(* IEC 61131-3 sources: 2026_Projet_YGO_ExcavatriceDragage/CODE/SIMULATION/PLC_TESTS, 3 files *)

(* ---- GVL_PLC_Tests.st ---- *)
(* ═══════════════════════════════════════════════════════════════
   🧪 GVL_PLC_Tests — Variables globales du banc de validation
   ───────────────────────────────────────────────────────────────
   🎯 Rôle : Regroupe toutes les commandes et retours d'états
      du banc de tests automatique in-PLC.
   ═══════════════════════════════════════════════════════════════ *)

{attribute 'qualified_only'}
VAR_GLOBAL
    CmdRunTests                : BOOL := FALSE; // 🔑 Lancement des tests de validation (bouton IHM/Simu)
    TestInProgress             : BOOL;          // Test en cours d'exécution
    AllTestsPassed             : BOOL;          // Succès global : tous les scénarios validés 🟢
    TestFailed                 : BOOL;          // Échec détecté 🔴
    TC01_NominalArming_Ok      : BOOL;          // Statut TC-01 (Armement nominal & AU)
    TC02_RedundancyFault_Ok    : BOOL;          // Statut TC-02 (Contacteur collé)
    TC03_Lockout_Ok            : BOOL;          // Statut TC-03 (Lockout 5s)
    FailedTestCase             : INT;           // Index du scénario en échec

    // Signaux de surcharge internes (pilotés par le validateur de test)
    OverrideChainTrue          : BOOL;          // Force la boucle AU à TRUE
    OverrideChainFalse         : BOOL;          // Force la boucle AU à FALSE
    OverrideContactorFalse     : BOOL;          // Force le retour contacteur à FALSE
END_VAR

(* ---- FB_PLC_Tests_Management.st ---- *)
(* ═══════════════════════════════════════════════════════════════
   🧪 FB_PLC_Tests_Management — Gestion Globale des Tests de Validation Automatisés
   ───────────────────────────────────────────────────────────────
   🎯 Rôle : Regroupe, configure et orchestre toutes les instances
      de tests de validation automate (banc de test global).
      Met à jour directement GVL_PLC_Tests pour affichage unifié.
   ═══════════════════════════════════════════════════════════════ *)

FUNCTION_BLOCK PUBLIC FB_PLC_Tests_Management
VAR
    // 🧱 Instances de tests individuels hébergées
    instSafetyValidation       : FB_SafetyValidation;

    // Flag de déclenchement interne
    TriggerSafetyTests         : BOOL;
END_VAR

// === IMPLEMENTATION ===

// 1. Détection du bit de déclenchement global dans GVL_PLC_Tests
IF GVL_PLC_Tests.CmdRunTests THEN
    GVL_PLC_Tests.CmdRunTests := FALSE;
    TriggerSafetyTests := TRUE;
ELSE
    TriggerSafetyTests := FALSE;
END_IF;

// 2. Appel de l'instance de test pour la sécurité d'urgence
instSafetyValidation(StartTests := TriggerSafetyTests);

// 3. Centralisation directe des résultats dans GVL_PLC_Tests
GVL_PLC_Tests.TestInProgress          := instSafetyValidation.TestInProgress;
GVL_PLC_Tests.AllTestsPassed          := instSafetyValidation.AllTestsPassed;
GVL_PLC_Tests.TestFailed              := instSafetyValidation.TestFailed;
GVL_PLC_Tests.TC01_NominalArming_Ok   := instSafetyValidation.TC01_NominalArming_Ok;
GVL_PLC_Tests.TC02_RedundancyFault_Ok := instSafetyValidation.TC02_RedundancyFault_Ok;
GVL_PLC_Tests.TC03_Lockout_Ok         := instSafetyValidation.TC03_Lockout_Ok;
GVL_PLC_Tests.FailedTestCase          := instSafetyValidation.FailedTestCase;

// 4. Centralisation directe des surcharges de simulation (overrides)
GVL_PLC_Tests.OverrideChainTrue       := instSafetyValidation.OverrideChainTrue;
GVL_PLC_Tests.OverrideChainFalse      := instSafetyValidation.OverrideChainFalse;
GVL_PLC_Tests.OverrideContactorFalse  := instSafetyValidation.OverrideContactorFalse;

(* ---- FB_SafetyValidation.st ---- *)
(* ═══════════════════════════════════════════════════════════════
   🧪 FB_SafetyValidation — Validateur Automatique de Sécurité
   ───────────────────────────────────────────────────────────────
   🎯 Rôle : Séquenceur de test sous forme de bloc fonctionnel (FB).
      Exécute les cas de tests réglementaires de la boucle d'urgence.
      En cas d'échec sur un test, passe au suivant pour tout valider.
      Résistant aux verrouillages temporels (Lockout 5s) entre tests.
   ═══════════════════════════════════════════════════════════════ *)

FUNCTION_BLOCK PUBLIC FB_SafetyValidation
VAR_INPUT
    StartTests                 : BOOL;        // Commande de démarrage des tests
END_VAR
VAR_OUTPUT
    // Rapport de test
    TestInProgress             : BOOL;
    TC01_NominalArming_Ok      : BOOL;
    TC02_RedundancyFault_Ok    : BOOL;
    TC03_Lockout_Ok            : BOOL;
    AllTestsPassed             : BOOL;
    TestFailed                 : BOOL;
    FailedTestCase             : INT;         // Index du scénario ayant échoué

    // Demandes de surcharge (overrides) vers le programme de simulation
    OverrideChainTrue          : BOOL;        // Force l'entrée boucle d'urgence à TRUE
    OverrideChainFalse         : BOOL;        // Force l'entrée boucle d'urgence à FALSE
    OverrideContactorFalse     : BOOL;        // Force l'entrée contacteur à FALSE
END_VAR
VAR
    StartTestEdge              : R_TRIG;
    TestSeqStep                : INT := 0;    // Séquenceur de test
    LastStep                   : INT := 0;    // Mémoire de l'étape précédente
    TestTimer                  : TON;         // Timer d'attente d'étapes (timeout)

    // Signaux locaux pour stimuler le bloc sous test
    ArmRequest                 : BOOL;
    ResetFaults                : BOOL;
    CmdEmergencyCutOff         : BOOL;
END_VAR

// === IMPLEMENTATION ===

// ⛔ Neutralisation si la simulation globale n'est pas active (sécurité physique)
IF NOT GVL_Simulation.SimulationModeActive THEN
    TestSeqStep := 0;
    TestInProgress := FALSE;
    OverrideChainTrue := FALSE;
    OverrideChainFalse := FALSE;
    OverrideContactorFalse := FALSE;
    RETURN;
END_IF;

StartTestEdge(CLK := StartTests);

// 🔄 Réinitialisation du timer d'étape si changement d'étape détecté
IF TestSeqStep <> LastStep THEN
    TestTimer(IN := FALSE);
    LastStep := TestSeqStep;
END_IF;

// ⏱️ Timer général d'étape (timeout de 10s maximum par étape)
TestTimer(IN := (TestSeqStep <> 0), PT := T#10s);

// 🚨 Échec automatique si le timer d'étape expire (sécurité anti-blocage)
IF TestTimer.Q AND TestSeqStep <> 0 AND TestSeqStep <> 999 THEN
    TestFailed := TRUE;

    // Si timeout dans TC-01 (étapes 10 à 17), on passe au TC-02 (étape 20)
    IF TestSeqStep >= 10 AND TestSeqStep <= 17 THEN
        OverrideChainFalse := FALSE;
        FailedTestCase := 1;
        TestSeqStep := 20;

    // Si timeout dans TC-02 (étapes 20 à 22), on passe au TC-03 (étape 30)
    ELSIF TestSeqStep >= 20 AND TestSeqStep <= 22 THEN
        OverrideChainTrue := FALSE;
        FailedTestCase := 2;
        TestSeqStep := 30;

    // Si timeout dans TC-03 (étapes 30 à 36), fin de séquence (étape 999)
    ELSE
        OverrideContactorFalse := FALSE;
        FailedTestCase := 3;
        TestSeqStep := 999;
    END_IF;
END_IF;

// 🔀 Séquenceur de Test Automatique
CASE TestSeqStep OF

    0: // IDLE — En attente du départ de test
        IF StartTestEdge.Q THEN
            TestInProgress := TRUE;
            TC01_NominalArming_Ok := FALSE;
            TC02_RedundancyFault_Ok := FALSE;
            TC03_Lockout_Ok := FALSE;
            AllTestsPassed := FALSE;
            TestFailed := FALSE;
            FailedTestCase := 0;
            OverrideChainTrue := FALSE;
            OverrideChainFalse := FALSE;
            OverrideContactorFalse := FALSE;
            TestSeqStep := 10;
        END_IF;

    // ─────────────────────────────────────────────────────────────────
    // 🧪 SCÉNARIO 1 : Séquence Nominale (TC-01)
    // ─────────────────────────────────────────────────────────────────
    10: // Phase 1.1 : Initialisation saine (attente fin du verrouillage de sécurité précédent)
        ResetFaults := TRUE;
        IF NOT PRG_10_Outputs.instSafetyEmergencyManagement.RedundancyTestFailed AND
           NOT PRG_10_Outputs.instSafetyEmergencyManagement.EmergencyArmingFailed AND
           NOT PRG_10_Outputs.instSafetyEmergencyManagement.EmergencyArmingLockoutActive THEN
            ResetFaults := FALSE;
            ArmRequest := TRUE; // Maintient la demande jusqu'au démarrage réel
            TestSeqStep := 11;
        END_IF;

    11: // Phase 1.2 : Envoi demande réarmement et attente début auto-test
        IF PRG_10_Outputs.instSafetyEmergencyManagement.ArmingSeqStep = 1 THEN
            ArmRequest := FALSE; // Relâche la demande
            TestSeqStep := 13;
        END_IF;

    13: // Phase 1.4 : Attente réussite de l'auto-test et début impulsion armement
        IF PRG_10_Outputs.instSafetyEmergencyManagement.ArmingSeqStep = 5 THEN
            TestSeqStep := 14;
        END_IF;

    14: // Phase 1.5 : Attente fin de l'impulsion et confirmation armement
        IF PRG_00_Inputs.EmergencyStopOk AND PRG_10_Outputs.instSafetyEmergencyManagement.ArmingSeqStep = 0 THEN
            // Armé nominalement ! Maintenant on teste le Trip d'urgence
            TestSeqStep := 15;
        END_IF;

    15: // Phase 1.6 : Simulation d'un appui bouton d'urgence (Coupure franche)
        OverrideChainFalse := TRUE;
        TestSeqStep := 16;

    16: // Phase 1.7 : Vérification coupure instantanée
        IF NOT PowerCutOff_A_RQ AND NOT PowerCutOff_B_RQ AND NOT PRG_00_Inputs.EmergencyStopOk THEN
            // Coupure validée, on relâche le bouton d'urgence (doit rester coupé)
            OverrideChainFalse := FALSE;
            TestSeqStep := 17;
        END_IF;

    17: // Phase 1.8 : Vérification de l'auto-maintien (Latch)
        IF NOT PowerCutOff_A_RQ AND NOT PowerCutOff_B_RQ THEN
            TC01_NominalArming_Ok := TRUE;
            TestSeqStep := 20; // Passer au test de redondance
        ELSE
            TestFailed := TRUE;
            FailedTestCase := 1;
            TestSeqStep := 20; // continue au test suivant
        END_IF;

    // ─────────────────────────────────────────────────────────────────
    // 🧪 SCÉNARIO 2 : Défaut de Redondance (TC-02)
    // ─────────────────────────────────────────────────────────────────
    20: // Phase 2.1 : Acquitter le défaut précédent et attendre la fin du verrouillage de sécurité
        ResetFaults := TRUE;
        IF NOT PRG_10_Outputs.instSafetyEmergencyManagement.RedundancyTestFailed AND
           NOT PRG_10_Outputs.instSafetyEmergencyManagement.EmergencyArmingLockoutActive THEN
            ResetFaults := FALSE;
            ArmRequest := TRUE; // Maintient la demande
            TestSeqStep := 21;
        END_IF;

    21: // Phase 2.2 : Attente de l'auto-test canal A
        IF PRG_10_Outputs.instSafetyEmergencyManagement.ArmingSeqStep = 1 THEN
            ArmRequest := FALSE; // Relâche la demande
            // Simuler contacteur A soudé
            OverrideChainTrue := TRUE;
            TestSeqStep := 22;
        END_IF;

    22: // Phase 2.3 : Vérification de la détection du défaut (dans les 200ms)
        IF PRG_10_Outputs.instSafetyEmergencyManagement.RedundancyTestFailed AND
           PRG_10_Outputs.instSafetyEmergencyManagement.ArmingSeqStep = 0 THEN
            // Détection réussie ! Les sorties doivent être inhibées.
            OverrideChainTrue := FALSE;
            TC02_RedundancyFault_Ok := TRUE;
            TestSeqStep := 30; // Passer au test de Lockout
        END_IF;

    // ─────────────────────────────────────────────────────────────────
    // 🧪 SCÉNARIO 3 : Verrouillage temporel (TC-03)
    // ─────────────────────────────────────────────────────────────────
    30: // Phase 3.1 : Acquitter et attendre la fin du verrouillage précédent
        ResetFaults := TRUE;
        IF NOT PRG_10_Outputs.instSafetyEmergencyManagement.RedundancyTestFailed AND
           NOT PRG_10_Outputs.instSafetyEmergencyManagement.EmergencyArmingLockoutActive THEN
            ResetFaults := FALSE;
            ArmRequest := TRUE; // Maintient la demande
            // Bloquer le contacteur de puissance à FALSE
            OverrideContactorFalse := TRUE;
            TestSeqStep := 31;
        END_IF;

    31: // Phase 3.2 : Attente du début d'auto-test pour relâcher le bouton
        IF PRG_10_Outputs.instSafetyEmergencyManagement.ArmingSeqStep = 1 THEN
            ArmRequest := FALSE;
        END_IF;
        IF PRG_10_Outputs.instSafetyEmergencyManagement.EmergencyArmingFailed AND
           PRG_10_Outputs.instSafetyEmergencyManagement.EmergencyArmingLockoutActive THEN
            TestSeqStep := 32;
        END_IF;

    32: // Phase 3.3 : Tenter de réarmer immédiatement pendant le lockout de 5s
        ArmRequest := TRUE;
        TestSeqStep := 33;

    33: // Phase 3.4 : Vérifier que la demande de réarmement est ignorée
        ArmRequest := FALSE;
        IF PRG_10_Outputs.instSafetyEmergencyManagement.ArmingSeqStep <> 0 THEN
            // Pas normal, on a démarré pendant le lockout !
            OverrideContactorFalse := FALSE;
            TestFailed := TRUE;
            FailedTestCase := 3;
            TestSeqStep := 999;
        ELSE
            // Demande ignorée avec succès, on attend la fin du lockout
            TestSeqStep := 34;
        END_IF;

    34: // Phase 3.5 : Attente de la libération du verrouillage (5s)
        IF NOT PRG_10_Outputs.instSafetyEmergencyManagement.EmergencyArmingLockoutActive THEN
            // Lockout terminé, on désactive le blocage contacteur
            OverrideContactorFalse := FALSE;
            ResetFaults := TRUE;
            TestSeqStep := 35;
        END_IF;

    35: // Phase 3.6 : Valider qu'un réarmement normal est à nouveau possible
        ResetFaults := FALSE;
        ArmRequest := TRUE;
        TestSeqStep := 36;

    36: // Phase 3.7 : Confirmation finale de l'armement après lockout
        IF PRG_10_Outputs.instSafetyEmergencyManagement.ArmingSeqStep = 1 THEN
            ArmRequest := FALSE;
        END_IF;
        IF PRG_00_Inputs.EmergencyStopOk THEN
            TC03_Lockout_Ok := TRUE;
            AllTestsPassed := NOT TestFailed; // Succès global si aucun échec intermédiaire
            TestSeqStep := 100; // Succès global !
        END_IF;

    100: // FIN DE CYCLE DE TEST (SUCCÈS OU ÉCHEC PARTIEL)
        TestInProgress := FALSE;
        TestSeqStep := 0;

    999: // ÉCHEC CRITIQUE / ABANDON
        TestInProgress := FALSE;
        TestSeqStep := 0;

END_CASE;

// === LIAISON DES ESTIMULI AUX VARIABLES D'ÉCHANGE GLOBALES ===
IF TestInProgress THEN
    GVL_IHM.Modes.CmdEmergencyArming := ArmRequest;
    GVL_IHM.Modes.FaultMachineReset  := ResetFaults;
END_IF;
